// TIA Portal V20 export
// export: Created 2026-10-12T16:46:22.8991769Z, ExportSetting WithDefaults, DisplayName Totally Integrated Automation Portal, DisplayVersion V20 Update 6, DisplayName TIA Portal Openness, DisplayVersion V20 Update 6, DisplayName TIA Portal Version Control Interface, DisplayVersion V20 Update 6, DisplayName SINAMICS Startdrive Advanced, DisplayVersion V20 SP1 Update 2, DisplayName SINAMICS Startdrive G110M, G120, G120C, G120D, G120P, G115D, DisplayVersion V20 SP1 Update 2, DisplayName SINAMICS Startdrive G130, G150, S120, S150, SINAMICS MV, G220, S200, S210, DisplayVersion V20 SP1 Update 2, DisplayName STEP 7 Professional, DisplayVersion V20 Update 6, DisplayName STEP 7 Safety, DisplayVersion V20 Update 2, DisplayName WinCC Basic/Comfort/Advanced, DisplayVersion V20 Update 6, DisplayName WinCC Professional, DisplayVersion V20 Update 6, DisplayName WinCC Unified, DisplayVersion V20 Update 6
TYPE "UDT_Badschritt"
// ==========================================================================
//  Badlogik Chemisch Nickel - Gesamtquelle v0.9
// 
//  Aenderungen v0.9:
//    - Pumpe_FU (Umwaelzpumpe Bad 25): Sollwert, Netzschuetz, Freigabe, Reset
//    - FU-Resets (WB1, WB2, Pumpe) im Handbetrieb steuerbar
//    - "Pumpe Bad 25(1)" entfernt (Relikt)
//    - "Motorschutz 275aQ1" und "Wartungsschalter (1)" entfernt (Relikt)
//    - FU-Steuerwerte in Rueckmeldung
//    - Tag-Aenderung: A0.6 = "Netzschuetz Pumpe Bad 25" (war "Pumpe Bad 25")
//    - Neue Tags: "FU Pumpe Freigabe" A4.5, "Reset FU Pumpe" A4.6,
//                 "Pumpen_FU_Steuerwert" QW64, "FU Pumpe bereit" E0.7
//    - Auftrag_Abgeschlossen[0..9] im DB_CPU_to_IPC (Handshake fuer IPC)
// ==========================================================================
// stored: IsFailsafeCompliant false
   STRUCT
      BadNr : Int;
      Verweilzeit : Time;
      Vorwarnzeit : Time;
      Kritische_Zeit : Time;
      Pumpe : Bool;
      Pumpe_FU_Soll : Real;   // Umwaelzpumpe Drehzahl (%)
      Ultraschall : Bool;
      Heizung : Real;
      Heizung_Toleranz : Real;
      Warenbewegung_X : Real;
      Warenbewegung_Y : Real;
      GR_Aktiv : Bool;
      GR_Strom_Soll : Real;
      GR_Spannung_Soll : Real;
      GR_Pulsfrequenz : Real;
      GR_DutyCycle : Real;
      Alarm_Aktiv : Bool;
   END_STRUCT;
END_TYPE
